Fanuc KAREL source: KT00607.KL

PROGRAM KT00607
%NOLOCKGROUP
VAR
  R1: REAL
  R2: REAL
  OUT: INTEGER
BEGIN
  R1 = 2.0
  R2 = 3.0
  R1 = 2.0
  R2 = 3.0
  OUT = NOT R1
END KT00607
